TYPE ST_Production_Parameter :
STRUCT
	
	stRecipe	: ST_Prod_Recipe;
	WeightOrder	: REAL;//kg
	arrWeightIng: ARRAY[1..g_Prod.cMaxCompInProduct] OF REAL;
	prodDT		: DT;
	prodDate	: DATE;
	prodTime	: TIME;
	
	timeRemainToStart: TIME;
	timeProductionDuration: TIME;
	
	eStatus		: E_Prod_Status;


	
	hmiRecipeIndex: INT;
	
	bGetRecipe	: BOOL;
	listRecipe	: ARRAY[1..g_Prod.cMax_Prod_Recipe] OF STRING(30);



END_STRUCT
END_TYPE

(* stored: Version 1.1.0.1, ProductVersion 3.1.4024.15
   DUT ST_Production_Parameter: Id {a644b6ea-1ad6-4088-8a4e-dec51479ebd2} *)
